FUNCTION_BLOCK F_MUX_16 (* multiplexer *)
  (* Standard: 61131-3; Classification: standard selection function; Description: Copyright (c) 2026 Meisterschulen am Ostbahnhof This program and the accompanying materials are made available under the terms of the Eclipse Public License 2.0 which is available at https://www.eclipse.org/legal/epl-2.0/ SPDX-License-Identifier: EPL-2.0 *)
  (* Version 1.0, 2026-10-11, Franz Höpfinger, Meisterschulen am Ostbahnhof, created from F_MUX_32 *)
  PACKAGE iec61131::selection;
  {SET_ATTRIBUTE(eclipse4diac::core::GenericClassName, 'GEN_F_MUX')}
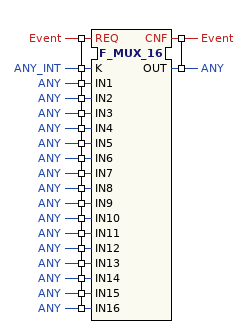
  EVENT_INPUT
    REQ WITH IN1, IN2, IN3, IN4, IN5, IN6, IN7, IN8, IN9, IN10, IN11, IN12, IN13, IN14, IN15, IN16, K; (* Service Request *)
  END_EVENT
  EVENT_OUTPUT
    CNF WITH OUT; (* Confirmation of Requested Service *)
  END_EVENT
  VAR_INPUT
    K : ANY_INT; (* Select one of n inputs *)
    IN1 : ANY; (* Input value 1 *)
    IN2 : ANY; (* Input value 2 *)
    IN3 : ANY; (* Input value 3 *)
    IN4 : ANY; (* Input value 4 *)
    IN5 : ANY; (* Input value 5 *)
    IN6 : ANY; (* Input value 6 *)
    IN7 : ANY; (* Input value 7 *)
    IN8 : ANY; (* Input value 8 *)
    IN9 : ANY; (* Input value 9 *)
    IN10 : ANY; (* Input value 10 *)
    IN11 : ANY; (* Input value 11 *)
    IN12 : ANY; (* Input value 12 *)
    IN13 : ANY; (* Input value 13 *)
    IN14 : ANY; (* Input value 14 *)
    IN15 : ANY; (* Input value 15 *)
    IN16 : ANY; (* Input value 16 *)
  END_VAR
  VAR_OUTPUT
    OUT : ANY; (* IN1 for K = 0, IN2 for K = 1, IN3 for K = 2, IN4 for K = 3, IN5 for K = 4, IN6 for K = 5, IN7 for K = 6, IN8 for K = 7, IN9 for K = 8, IN10 for K = 9, IN11 for K = 10, IN12 for K = 11, IN13 for K = 12, IN14 for K = 13, IN15 for K = 14, IN16 for K = 15 *)
  END_VAR
END_FUNCTION_BLOCK
